Staubli VAL3: setBaseJOG.pgx

public program setBaseJOG(num x_nIndexTool)
  local tool l_tTool
  local frame l_fFrame
begin

  call getTool(x_nIndexTool,tMTool)
  //call getFrame(x_nIndexFrame,fMFrame)

  $jogContext(tMTool,world,0)
  logMsg("setMovePara:tool"+toString("",x_nIndexTool))
end
